(* IEC 61131-3 sources: Motor-Speed-Control-PLC-FPGA/PLC, 5 files *)

(* ---- GVL_MODBUS.iecst ---- *)
VAR_GLOBAL
    g_iPWM AT %MW0 : INT := 0;
    g_iSetpoint AT %MW1 : INT := 0;
    g_iDirection AT %MW2 : INT := 0;
END_VAR

(* ---- MODBUS.iecst ---- *)
PROGRAM MODBUS
VAR
    xSW1 : BOOL AT %IX0.2;
    xSW2 : BOOL AT %IX0.3;
    xSW3 : BOOL AT %IX0.4;
    xSW4 : BOOL AT %IX0.5;
    xSW5 : BOOL AT %IX0.6;
    xSW6 : BOOL AT %IX0.7;
    xSW7 : BOOL AT %IX0.8;

    xDirectionSwitch : BOOL AT %IX0.9;
    iSetpointTemp : INT := 0;
END_VAR

iSetpointTemp := 0;

IF xSW1 THEN iSetpointTemp := iSetpointTemp + 1; END_IF;
IF xSW2 THEN iSetpointTemp := iSetpointTemp + 2; END_IF;
IF xSW3 THEN iSetpointTemp := iSetpointTemp + 4; END_IF;
IF xSW4 THEN iSetpointTemp := iSetpointTemp + 8; END_IF;
IF xSW5 THEN iSetpointTemp := iSetpointTemp + 16; END_IF;
IF xSW6 THEN iSetpointTemp := iSetpointTemp + 32; END_IF;
IF xSW7 THEN iSetpointTemp := iSetpointTemp + 64; END_IF;

GVL_MODBUS.g_iSetpoint := iSetpointTemp;

IF xDirectionSwitch THEN
    GVL_MODBUS.g_iDirection := 1;
ELSE
    GVL_MODBUS.g_iDirection := 0;
END_IF;

(* ---- PRG_HSC.iecst ---- *)
PROGRAM PRG_HSC
VAR
    xHSCInitDone : BOOL := FALSE;
    xSyncPulse : BOOL := FALSE;

    udiCount0 : UDINT := 0;
    udiCount1 : UDINT := 0;

    xValid0 : BOOL := FALSE;
    xValid1 : BOOL := FALSE;
    xError0 : BOOL := FALSE;
    xError1 : BOOL := FALSE;
END_VAR

IF NOT xHSCInitDone THEN
    xSyncPulse := TRUE;
    xHSCInitDone := TRUE;
ELSE
    xSyncPulse := FALSE;
END_IF;

HSC_Forward(
    Enable := TRUE,
    Sync := xSyncPulse,
    ACK_Modulo := FALSE
);

HSC_Reverse(
    Enable := TRUE,
    Sync := xSyncPulse,
    ACK_Modulo := FALSE
);

xValid0 := HSC_Forward.Validity;
xError0 := HSC_Forward.Error;
IF xValid0 THEN
    udiCount0 := DWORD_TO_UDINT(HSC_Forward.CurrentValue);
END_IF;

xValid1 := HSC_Reverse.Validity;
xError1 := HSC_Reverse.Error;
IF xValid1 THEN
    udiCount1 := DWORD_TO_UDINT(HSC_Reverse.CurrentValue);
END_IF;

(* ---- PRG_PID.iecst ---- *)
PROGRAM PRG_PID

VAR

     (* FALSE хэвээр эхэлнэ. Онлайн monitor-оор TRUE болгож PID-ийг идэвхжүүлнэ. *)
    xPID_Enable : BOOL :=TRUE;

    rSetpointRPM : REAL := 0.0;
    rActualRPM : REAL := 0.0;
    rError : REAL := 0.0;
    rPreviousError : REAL := 0.0;

    (* Эхний туршилтын коэффициентууд. Бодит мотор дээр тохируулна. *)
    rKp : REAL := 0.50;
    rKi : REAL := 0.05;
    rKd : REAL := 0.0;

    rP : REAL := 0.0;
    rI : REAL := 0.0;
    rD : REAL := 0.0;
    rIntegral : REAL := 0.0;

    rRawOutput : REAL := 0.0;
    rPWM : REAL := 0.0;
    rTs : REAL := 0.5;

    uiPWM_Command : UINT := 0;
    xFirstPIDSample : BOOL := TRUE;

END_VAR

xPID_Enable := TRUE;

(* RPM шинэ sample гарсан үед л PID тооцно *)
IF PRG_RPM.xSampleTick THEN

    IF xPID_Enable THEN
        (* Setpoint нь MW1-ээс уншигдана *)
        rSetpointRPM := INT_TO_REAL(GVL_MODBUS.g_iSetpoint);

        (* Direction=0 бол sensor 0, Direction=1 бол sensor 1-ийн RPM *)
        IF GVL_MODBUS.g_iDirection = 0 THEN
            rActualRPM := PRG_RPM.rRPM0;
        ELSE
            rActualRPM := PRG_RPM.rRPM1;
        END_IF;

        IF rSetpointRPM <= 0.0 THEN
            rPWM := 0.0;
            uiPWM_Command := 0;
            rIntegral := 0.0;
            rPreviousError := 0.0;
            rP := 0.0;
            rI := 0.0;
            rD := 0.0;
            xFirstPIDSample := TRUE;

        ELSE
            (* Алдаа: зорилтот хурд - бодит хурд *)
            rError := rSetpointRPM - rActualRPM;

            (* Proportional *)
            rP := rKp * rError;

            (* Derivative. Эхний sample дээр 0 *)
            IF xFirstPIDSample THEN
                rD := 0.0;
                xFirstPIDSample := FALSE;
            ELSE
                rD := rKd * (rError - rPreviousError) / rTs;
            END_IF;

            (* Өмнөх integral-тай түр гаралт бодож anti-windup шийдэх *)
            rI := rKi * rIntegral;
            rRawOutput := rP + rI + rD;

            (* Гаралт saturation-д хүрээгүй, эсвэл saturation-аас буцах
               чиглэлийн алдаа гарсан үед л integral-ийг нэмнэ *)
            IF ((rRawOutput < 255.0) AND (rRawOutput > 0.0)) OR
               ((rRawOutput >= 255.0) AND (rError < 0.0)) OR
               ((rRawOutput <= 0.0) AND (rError > 0.0)) THEN
                rIntegral := rIntegral + (rError * rTs);
            END_IF;

            (* Integral хуримтлалыг хязгаарлах *)
            IF rIntegral > 1000.0 THEN
                rIntegral := 1000.0;
            ELSIF rIntegral < -1000.0 THEN
                rIntegral := -1000.0;
            END_IF;

            (* PID-ийн нийлбэр гаралт *)
            rI := rKi * rIntegral;
            rRawOutput := rP + rI + rD;

            (* PWM команд 0..255 хүрээнд хязгаарлах *)
            IF rRawOutput > 255.0 THEN
                rPWM := 255.0;
            ELSIF rRawOutput < 0.0 THEN
                rPWM := 0.0;
            ELSE
                rPWM := rRawOutput;
            END_IF;

            uiPWM_Command := REAL_TO_UINT(rPWM);
            rPreviousError := rError;
        END_IF;

    ELSE
        (* PID disabled үед PWM=0 *)
        rPWM := 0.0;
        uiPWM_Command := 0;
        rIntegral := 0.0;
        rPreviousError := 0.0;
        rP := 0.0;
        rI := 0.0;
        rD := 0.0;
        xFirstPIDSample := TRUE;
    END_IF;
  (* PWM үр дүнг MW0-д бичнэ. FPGA зөвхөн энэ регистрийг уншина. *)
    GVL_MODBUS.g_iPWM := UINT_TO_INT(uiPWM_Command);
END_IF;

(* ---- PRG_RPM.iecst ---- *)
PROGRAM PRG_RPM
VAR
    tmSample : TON;
    xSampleTick : BOOL := FALSE;

    udiPPR0 : UDINT := 10;
    udiPPR1 : UDINT := 10;

    udiCount0 : UDINT := 0;
    udiCount1 : UDINT := 0;
    udiPrev0 : UDINT := 0;
    udiPrev1 : UDINT := 0;
    udiDelta0 : UDINT := 0;
    udiDelta1 : UDINT := 0;

    rRPM0 : REAL := 0.0;
    rRPM1 : REAL := 0.0;
END_VAR

tmSample(
    IN := NOT tmSample.Q,
    PT := T#500ms
);

xSampleTick := tmSample.Q;

IF xSampleTick THEN
    udiCount0 := PRG_HSC.udiCount0;
    udiCount1 := PRG_HSC.udiCount1;

    IF udiCount0 >= udiPrev0 THEN
        udiDelta0 := udiCount0 - udiPrev0;
    ELSE
        udiDelta0 := 0;
    END_IF;

    IF udiCount1 >= udiPrev1 THEN
        udiDelta1 := udiCount1 - udiPrev1;
    ELSE
        udiDelta1 := 0;
    END_IF;

    udiPrev0 := udiCount0;
    udiPrev1 := udiCount1;

    IF udiPPR0 > 0 THEN
        rRPM0 := UDINT_TO_REAL(udiDelta0) * 120.0 / UDINT_TO_REAL(udiPPR0);
    ELSE
        rRPM0 := 0.0;
    END_IF;

    IF udiPPR1 > 0 THEN
        rRPM1 := UDINT_TO_REAL(udiDelta1) * 120.0 / UDINT_TO_REAL(udiPPR1);
    ELSE
        rRPM1 := 0.0;
    END_IF;
END_IF;
